{attribute 'no_assign'}
FUNCTION_BLOCK FB_DO_WTURBINE_LD0_WTUR1_TotWh EXTENDS FB_AcsiCommonDataClass
VAR_INPUT
	cntVal: FB_DO_WTURBINE_LD0_WTUR1_TotWh_cntVal := (sClass:='BCR', bLinkResult:=THIS^.AddDataToContainer(ipData:=cntVal));
END_VAR
VAR
END_VAR

END_FUNCTION_BLOCK

(* stored: Version 1.1.0.1
   POU FB_DO_WTURBINE_LD0_WTUR1_TotWh: Id {a0cfac60-ee05-45be-b7ac-62e3ca9bc5ed}, SpecialFunc None *)
